Staubli VAL3: MoveJ.pgx

public program MoveJ(jointRx x_jPoint, tool x_tTool, mdesc x_mSpeed, num& x_nMoveId, bool x_bExact)
// // 关节运动movej程序
// // 用该程序替代原val3程序中的movej()指令即可
// // 因为原move指令有返回值moveID，所以这里引入一个x_nMoveId，随参考传递出来
  local bool l_bResult
begin
  // ---------------------------------------------------------------------------- //
  // 关节运动movej程序
  // 用该程序替代原val3程序中的movej()指令即可
  // 因为原move指令有返回值moveID，所以这里引入一个x_nMoveId，随参考传递出来
  // ---------------------------------------------------------------------------- //
  //
  //
  l_bResult=isInRange(x_jPoint)
  if l_bResult==true
    x_nMoveId=movej(x_jPoint,x_tTool,x_mSpeed)
    if x_bExact
      waitEndMove()
    endIf
    // log
    call logMoveMsgJ(x_jPoint,x_tTool,x_mSpeed,x_nMoveId,x_bExact)
  else
    // 关节点位超限
  endIf

end
